Fanuc KAREL source: KO00067.KL

PROGRAM KO00067
%NOLOCKGROUP
%ENVIRONMENT MIR
VAR
  P1: XYZWPREXT
  P2: POSITION
  F: BOOLEAN
  OUT: XYZWPREXT
BEGIN
  F = TRUE
  OUT = MIRROR(P1, P2, F)
END KO00067
